TYPE "ST_UserRecord"
VERSION : 0.1
   STRUCT
      User : String[32];
      Salt : Array[0..15] of Byte;
      PinHash : Array[0..31] of Byte;
      Level : DInt;
   END_STRUCT;

END_TYPE

